Fanuc KAREL source: kb00202.KL

-- PROVISIONAL review KL for V940-1; original PC SHA256 a6d81da5dc243b993e837b8ffc2028353ca0a724f761e9adbfd182254843eecd
-- Incomplete behavior may be omitted. Consult companion uncertainty JSON. Do not deploy.
PROGRAM KB00202
%NOLOCKGROUP
BEGIN
  -- V9_ZERO_TABLE_METADATA_HINT layout=0002_ascii; no indexed target words; source/name/runtime held
  -- UNRESOLVED_PC offsets 5-14; opcodes 3F,75
  -- UNRESOLVED_PC offsets 19-28; opcodes 3F,75
  -- UNRESOLVED_PC offsets 33-40; opcodes 9D,23
  -- UNRESOLVED_PC offsets 45-77; opcodes 27,22,22,2A,22,2A,22,31
  -- UNRESOLVED_PC offsets 82-86; opcodes 7F
END KB00202
